{attribute 'qualified_only'}
VAR_GLOBAL
	iContent_Main: INT;

END_VAR

(* stored: Version 1.1.0.1, ProductVersion 3.1.4024.13
   GVL g_Common: Id {d60cb8e0-5512-40e7-bb50-cbcec5ecabdd} *)
